PROGRAM MAIN
VAR
	// TcUnit finds every FB_TestSuite instance by itself; it is enough to declare them here.
	fbHomeDropReasonTests	: FB_HomeDropReason_Tests;
	fbHomeHoldTests			: FB_HomeHold_Tests;
	fbStartRequestTests		: FB_StartRequest_Tests;
	fbStepDrainTests		: FB_StepDrain_Tests;
	fbSweepStopTests		: FB_SweepStop_Tests;
	fbPointingForwardTests	: FB_PointingModelForward_Tests;
	fbIagRigTests			: FB_IagRig_Tests;
	fbStopDuringSlewTests	: IagStopDuringSlew_Tests;
	fbResetUnderMotionTests	: IagResetUnderMotion_Tests;
	fbErrorParkTests		: IagErrorPark_Tests;
	fbIagTimeoutsTests : IagTimeouts_Tests;
	fbParkDuringPowerOnTests	: IagParkDuringPowerOn_Tests;
	fbStopDuringParkTests	: IagStopDuringPark_Tests;
	fbParkInLimitTests		: IagParkInLimit_Tests;
	fbStuckStopTests		: IagStuckStop_Tests;
	fbCommandInputsTests	: IagCommandInputs_Tests;
	fbCommandAcceptanceTests	: IagCommandAcceptance_Tests;
	fbAbortStopTests		: IagAbortStop_Tests;
	fbParkPowerResetTests	: IagParkPowerReset_Tests;
	fbSupersedeTests		: IagSupersede_Tests;
	fbTelemetryTests		: IagTelemetry_Tests;
	fbCoordinatesTests		: IagCoordinates_Tests;
END_VAR

TcUnit.RUN();

END_PROGRAM

(* stored: Version 1.1.0.1, ProductVersion 3.1.4024.15
   POU MAIN: Id {8cc549e7-d335-44fc-af47-98df09911d71}, SpecialFunc None *)
